(* IEC 61131-3 sources: Test-Git_ESME26/TestProgettoESME_26.fbsproj/PacDriveLib Migration/Motion/Homing/PDL_FB_HomeSetPos.fb.st^, 3 files *)

(* ---- Init_Interfaces.meth.st ---- *)
METHOD PRIVATE Init_Interfaces : BOOL
VAR_INPUT
END_VAR

		Init_Interfaces := FALSE;

		IF
			i_etMode = PDL_ET_HomeSetPosMode.SetPosAxisAndLogEncoderPosition OR
			i_etMode = PDL_ET_HomeSetPosMode.RestorePosFromRetain OR
			i_etMode = PDL_ET_HomeSetPosMode.SetPosAxisPosition OR
			i_etMode = PDL_ET_HomeSetPosMode.RestorePosFromAxisencoder
		THEN
			IF i_ifDrive = 0 THEN
				SetDiagOutput(i_etDiag := GD.ET_Diag.InputParameterInvalid, i_etDiagExt := PDL_ET_DiagExt.DriveInvalid, i_sMsg := 'i_ifDrive = 0');
				diState := 0;
				RETURN;
			ELSE
				xSuccess := __QUERYINTERFACE(i_ifDrive, ifGetParentDevice);
				IF NOT xSuccess OR ifGetParentDevice = 0 THEN
					SetDiagOutput(
						i_etDiag    := GD.ET_Diag.InputParameterInvalid,
						i_etDiagExt := PDL_ET_DiagExt.DriveInvalid,
						i_sMsg      := 'i_ifDrive - IF_GetParentDevice not implemented.'
					);
					diState := 0;
					RETURN;
				END_IF

				ifDeviceAccess := ifGetParentDevice.GetParentDevice();

				xSuccess := __QUERYINTERFACE(ifDeviceAccess, ifScalingAccess);
				IF (NOT xSuccess OR ifScalingAccess = 0) THEN
					SetDiagOutput(
						i_etDiag    := GD.ET_Diag.InputParameterInvalid,
						i_etDiagExt := PDL_ET_DiagExt.DriveInvalid,
						i_sMsg      := 'i_ifDrive - IF_Scaling not implemented.'
					);
					diState := 0;
					RETURN;
				END_IF
				ifScaling := ifScalingAccess.Scaling;

				xSuccess := __QUERYINTERFACE(ifDeviceAccess, ifEncoderAccess);
				IF (NOT xSuccess OR ifEncoderAccess = 0) THEN
					SetDiagOutput(
						i_etDiag    := GD.ET_Diag.InputParameterInvalid,
						i_etDiagExt := PDL_ET_DiagExt.DriveInvalid,
						i_sMsg      := 'i_ifDrive - IF_Encoder not implemented.'
					);
					diState := 0;
					RETURN;
				END_IF
				ifEncoder := ifEncoderAccess.Encoder;

			END_IF
		END_IF

		IF i_etMode = PDL_ET_HomeSetPosMode.SetPosLogEncoderPosition OR i_etMode = PDL_ET_HomeSetPosMode.SetPosAxisAndLogEncoderPosition THEN
			IF iq_lencEncoder = 0 THEN
				SetDiagOutput(
					i_etDiag := GD.ET_Diag.InputParameterInvalid, i_etDiagExt := PDL_ET_DiagExt.LencInvalid, i_sMsg := 'iq_lencEncoder = 0'
				);
				diState := 0;
				RETURN;
			END_IF
		END_IF

		Init_Interfaces := TRUE;

(* ---- RegisterLoggerPoint.meth.st ---- *)
METHOD PUBLIC RegisterLoggerPoint
VAR_INPUT
	i_ifParent		: APL.IF_LoggerPoint;
	i_sName			: STRING[80];
END_VAR
VAR_OUTPUT
	q_etDiag		: GD.ET_Diag := GD.ET_Diag.Ok;
	q_etDiagExt		: PDL_ET_DiagExt := PDL_ET_DiagExt.Ok;
END_VAR
VAR
	etDiagBuffer		: GD.ET_Diag;
	etDiagExtBufferAPL	: APL.ET_DiagExt;
END_VAR

THIS^.fbLoggerPoint.RegisterLoggerPoint(	i_ifParent		:= i_ifParent,
											i_sName			:= i_sName,
											i_sType			:= 'FB_HomeSetPos',
											i_sSource		:= 'PDL',
											q_etDiag		=> etDiagBuffer,
											q_etDiagExt		=> etDiagExtBufferAPL);
IF (etDiagBuffer <> GD.ET_Diag.Ok) THEN
	CASE etDiagExtBufferAPL OF
		APL.ET_DiagExt.ParentInvalid:
			q_etDiag := GD.ET_Diag.InputParameterInvalid;
			q_etDiagExt := PDL_ET_DiagExt.ParentInvalid;

		APL.ET_DiagExt.ParentNotRegistered:
			q_etDiag := GD.ET_Diag.InputParameterInvalid;
			q_etDiagExt := PDL_ET_DiagExt.ParentNotRegistered;

		APL.ET_DiagExt.MaxNumberOfLoggerPointsExeeded:
			q_etDiag := GD.ET_Diag.InputParameterInvalid;
			q_etDiagExt := PDL_ET_DiagExt.MaxNumberOfLoggerPointsExeeded;

	ELSE
		q_etDiag := GD.ET_Diag.UnexpectedProgramBehavior;
		q_etdiagExt := PDL_ET_DiagExt.UnexpectedDiagExt;
	END_CASE
END_IF

(* ---- SetDiagOutput.meth.st ---- *)
METHOD PRIVATE SetDiagOutput : BOOL
VAR_INPUT
	i_etDiag	: GD.ET_Diag;
	i_etDiagExt	: PDL_ET_DiagExt;
	i_sMsg		: STRING[80];
END_VAR
VAR
END_VAR

IF i_etDiag <> GD.ET_Diag.Ok THEN
	q_xReady := FALSE;
END_IF
IF q_etDiag = GD.ET_Diag.OK OR i_etDiagExt = PDL_ET_DiagExt.Disabled THEN
	q_etDiag := i_etDiag;
	q_etDiagExt := i_etDiagExt;
	q_sMsg := i_sMsg;

	IF(i_etDiag = GD.ET_Diag.Ok) AND (THIS^.fbLoggerPoint.etLogLevel >= APL.ET_LogLevel.StatusMessage) THEN
		THIS^.fbLoggerPoint.AddLogEntry(	i_etLogLevel	:= APL.ET_LogLevel.StatusMessage,
											i_etDiag		:= q_etDiag,
											i_udiDiagExt	:= q_etDiagExt,
											i_sMessage		:= SE_CTBX.FC_MultiConcat(	i_sString1	:= Standard.CONCAT('ET_Diag: ', GD.FC_EtDiagToString(q_etDiag)),
																				i_sString2	:= Standard.CONCAT(' PDL_ET_DiagExt: ', PDL_FC_EtDiagExtToString(q_etDiagExt)),
																				i_sString3	:= Standard.CONCAT(' sMsg: ', q_sMsg),
																				i_sString4	:= ''),
											q_etDiag		:= ,	// ignore result
											q_etDiagExt		:= );	// ignore result
	ELSIF(i_etDiag = GD.ET_Diag.UnexpectedProgramBehavior) AND (THIS^.fbLoggerPoint.etLogLevel >= APL.ET_LogLevel.CriticalException) THEN
		THIS^.fbLoggerPoint.AddLogEntry(	i_etLogLevel	:= APL.ET_LogLevel.CriticalException,
											i_etDiag		:= q_etDiag,
											i_udiDiagExt	:= q_etDiagExt,
											i_sMessage		:= SE_CTBX.FC_MultiConcat(	i_sString1	:= Standard.CONCAT('ET_Diag: ', GD.FC_EtDiagToString(q_etDiag)),
																				i_sString2	:= Standard.CONCAT(' PDL_ET_DiagExt: ', PDL_FC_EtDiagExtToString(q_etDiagExt)),
																				i_sString3	:= Standard.CONCAT(' sMsg: ', q_sMsg),
																				i_sString4	:= ''),
											q_etDiag		:= ,	// ignore result
											q_etDiagExt		:= );	// ignore result
	ELSIF(i_etDiag <> GD.ET_Diag.Ok) AND (THIS^.fbLoggerPoint.etLogLevel >= APL.ET_LogLevel.Exception) THEN
		THIS^.fbLoggerPoint.AddLogEntry(	i_etLogLevel	:= APL.ET_LogLevel.Exception,
											i_etDiag		:= q_etDiag,
											i_udiDiagExt	:= q_etDiagExt,
											i_sMessage		:= SE_CTBX.FC_MultiConcat(	i_sString1	:= Standard.CONCAT('ET_Diag: ', GD.FC_EtDiagToString(q_etDiag)),
																				i_sString2	:= Standard.CONCAT(' PDL_ET_DiagExt: ', PDL_FC_EtDiagExtToString(q_etDiagExt)),
																				i_sString3	:= Standard.CONCAT(' sMsg: ', q_sMsg),
																				i_sString4	:= ''),
											q_etDiag		:= ,	// ignore result
											q_etDiagExt		:= );	// ignore result
	END_IF
END_IF
